(* IEC 61131-3 sources: avi-aoi-management/scripts/ai-eval/ngau-nhien/kho/st-ud4-may-tron-me/khung/src, 2 files *)

(* ---- KhoaLienDongVan.st ---- *)
FUNCTION_BLOCK KhoaLienDongVan
VAR_INPUT
    YC_A : BOOL;
    YC_B : BOOL;
    YC_XA : BOOL;
END_VAR
VAR_OUTPUT
    VAN_A : BOOL;
    VAN_B : BOOL;
    VAN_XA : BOOL;
    XUNG_DOT : BOOL;
END_VAR
    (* TODO: cài đặt theo đề bài *)
    VAN_A := FALSE;
END_FUNCTION_BLOCK

(* ---- MayTronMe.st ---- *)
FUNCTION_BLOCK MayTronMe
VAR_INPUT
    START : BOOL;
    STOP : BOOL;
    MUC : REAL;
    MUC_A : REAL;
    MUC_B : REAL;
    MUC_RONG : REAL;
    T_TRON : TIME;
END_VAR
VAR_OUTPUT
    VAN_A : BOOL;
    VAN_B : BOOL;
    VAN_XA : BOOL;
    MOTOR : BOOL;
    TRANG_THAI : INT;
    SO_ME : DINT;
END_VAR
    (* TODO: cài đặt theo đề bài *)
    VAN_A := FALSE;
END_FUNCTION_BLOCK
